(* IEC 61131-3 sources: veristc/veri-stc/tests/compiler-tests/negative, 18 files *)

(* ---- in_out_expr.st ---- *)
(* ================================================================
   negative/in_out_expr.st  --  VAR_IN_OUT 实参必须是简单变量名

   别名需要一个稳定的存储位置，表达式/常量没有地址可取，
   故 a1.ACC := SHARED + 1 必须被拒绝。
   ================================================================ *)

VAR_GLOBAL
  SHARED : DINT;
  a1 : ACCUM;
END_VAR

FUNCTION_BLOCK ACCUM
VAR_IN_OUT
  ACC : DINT;
END_VAR
  ACC := ACC + 1;
END_FUNCTION_BLOCK

PROGRAM MAIN
  a1(ACC := SHARED + 1);
END_PROGRAM

(* ---- in_out_local.st ---- *)
(* ================================================================
   negative/in_out_local.st  --  VAR_IN_OUT 别名目标不能是调用方局部

   MAIN 的 tick 是帧局部槽位（不在可寻址线性内存中），取不到地址，
   因此不能作为 a1.ACC 的别名目标。检查层必须以 alias 诊断拒绝。
   ================================================================ *)

VAR_GLOBAL
  a1 : ACCUM;
END_VAR

FUNCTION_BLOCK ACCUM
VAR_IN_OUT
  ACC : DINT;
END_VAR
  ACC := ACC + 1;
END_FUNCTION_BLOCK

PROGRAM MAIN
VAR
  tick : DINT;
END_VAR
  a1(ACC := tick);
END_PROGRAM

(* ---- in_out_type.st ---- *)
(* ================================================================
   negative/in_out_type.st  --  VAR_IN_OUT 两侧类型必须完全一致

   别名不经过隐式转换（同一块存储被两侧按同一宽度读写），
   且解引用指令按 4 字节定宽访问，故 INT(16 位) 目标必须拒绝。
   ================================================================ *)

VAR_GLOBAL
  SMALL : INT;
  a1 : ACCUM;
END_VAR

FUNCTION_BLOCK ACCUM
VAR_IN_OUT
  ACC : DINT;
END_VAR
  ACC := ACC + 1;
END_FUNCTION_BLOCK

PROGRAM MAIN
  a1(ACC := SMALL);
END_PROGRAM

(* ---- in_out_unbound.st ---- *)
(* ================================================================
   negative/in_out_unbound.st  --  VAR_IN_OUT 端口必须被绑定

   端口不绑定就没有别名目标（既无初值可拷贝，也无副本语义可言），
   与 IEC 要求一致：必须显式绑定到调用方存储。
   ================================================================ *)

VAR_GLOBAL
  SHARED : DINT;
  a1 : ACCUM;
END_VAR

FUNCTION_BLOCK ACCUM
VAR_IN_OUT
  ACC : DINT;
END_VAR
  ACC := ACC + 1;
END_FUNCTION_BLOCK

PROGRAM MAIN
  a1();
END_PROGRAM

(* ---- in_out_unknown_port.st ---- *)
(* ================================================================
   negative/in_out_unknown_port.st  --  调用只能绑定已声明端口

   FB_ACC 只声明了 ACC，调用点写 NOPE := SHARED 属于拼写/绕过声明，
   在逐引用端口上尤其危险（会把地址压进错误的槽位）。
   ================================================================ *)

VAR_GLOBAL
  SHARED : DINT;
  a1 : FB_ACC;
END_VAR

FUNCTION_BLOCK FB_ACC
VAR_IN_OUT
  ACC : DINT;
END_VAR
  ACC := ACC + 1;
END_FUNCTION_BLOCK

PROGRAM MAIN
  a1(ACC := SHARED, NOPE := SHARED);
END_PROGRAM

(* ---- literal_derived_name.st ---- *)
(* ================================================================
   negative/literal_derived_name.st -- 派生名不可书写

   expand_instances 产出的扁平全局名形如 a1#Q（'#' 为保留分隔符）。
   标识符文法是 字母 (字母|数字|_)*，不含 '#' ⇒ 源码里写 a1#Q 只能
   在词法阶段失败，用户无法伪造出一个"看起来像派生名"的名字去和
   真实派生名抢同一槽位，也不必再靠命名约定避免 a1_Q 这类碰撞。

   合法的字段访问写法是 IEC 点号 a1.Q，由 parser 融合为 a1#Q。
   ================================================================ *)

VAR_GLOBAL
  a1 : LATCH;
  x : DINT;
END_VAR

FUNCTION_BLOCK LATCH
VAR_OUTPUT
  Q : DINT;
END_VAR
  Q := 1;
END_FUNCTION_BLOCK

PROGRAM MAIN
  x := a1#Q;
END_PROGRAM

(* ---- name_collision_expanded.st ---- *)
(* ================================================================
   negative/name_collision_expanded.st -- 展开后派生名重复

   expand_instances（function_check.v）为实例 a1 的每个可写字段生成
   扁平全局名 a1#<字段>。若同一个 FUNCTION_BLOCK 里两个可写字段同名
   （此处 VAR_OUTPUT Q 与实例状态 VAR Q 重名），展开后就会产出两条
   a1#Q 声明 ⇒ 两个逻辑变量落到同一全局槽位、互相覆盖。

   这类冲突只在 prepare_program 之后才存在，因此 GATE-1 的重复名检查
   必须在展开后再跑一次，由 duplicate_declaration_msg 报出冲突的名字。

   （分隔符已改为标识符文法外的 '#'，用户无法手写派生名，所以静态
     命名冲突只剩"展开自身产出重名"这一条路径 —— 正是本用例。）
   ================================================================ *)

VAR_GLOBAL
  a1 : LATCH;
END_VAR

FUNCTION_BLOCK LATCH
VAR_INPUT
  K : DINT;
END_VAR
VAR_OUTPUT
  Q : DINT;
END_VAR
VAR
  Q : DINT;
END_VAR
  Q := K;
END_FUNCTION_BLOCK

PROGRAM MAIN
VAR
  tick : DINT;
END_VAR
  tick := CycleCounter();
  a1(K := tick);
END_PROGRAM

(* ---- qualified_in_out_read.st ---- *)
(* ================================================================
   negative/qualified_in_out_read.st -- 封装：别名端口不可用点号引用

   6.5.1 方向表的 VAR_IN_OUT 行。v1.5 起 VAR_IN_OUT 降级为"持有调用方
   存储地址的形参槽"（I32_LOAD_PTR / I32_STORE_PTR），expand_instances
   不为它生成派生全局，所以 `x := a1.ACC;` 引用的名字根本不存在，由类型
   检查阶段以 KIND=type 拒绝。

   这不是多余的严格性：调用方本来就持有别名目标（此处 shared），要读就
   直接读它 —— 读得到同一份存储，且不需要绕过 FB 的端口约定。

   与 qualified_input_read.st 的区别只在端口方向（IN_OUT vs INPUT）；
   与 qualified_internal_read.st（KIND=access）的区别在于名字是否存在。
   ================================================================ *)

(* 实例声明必须先于 POU 列表（顶层文法：VAR_GLOBAL → POU*）*)
VAR_GLOBAL
  a1 : ACCUM;
  shared : DINT;
  x : DINT;
END_VAR

FUNCTION_BLOCK ACCUM
VAR_INPUT
  K : DINT;
END_VAR
VAR_OUTPUT
  LAST : DINT;
END_VAR
VAR_IN_OUT
  ACC : DINT;
END_VAR
  LAST := ACC;
  ACC := ACC + K;
END_FUNCTION_BLOCK

PROGRAM MAIN
  a1(ACC := shared, K := 10);
  x := a1.ACC;
END_PROGRAM

(* ---- qualified_input_read.st ---- *)
(* ================================================================
   negative/qualified_input_read.st -- 封装：输入/别名端口不可用点号引用

   spec/safest-spec.md 6.5.1 方向表里 `VAR_INPUT` 与 `VAR_IN_OUT` 两行的
   体外访问都落到 `KIND=type`：expand_instances 只为可写字段
   （VAR_OUTPUT + 实例内 VAR）生成扁平派生全局，输入端口经调用点绑定为
   形参、别名端口降级为指针形参，二者都不存在名为 a1#K / a1#ACC 的全局。
   于是引用它们 = 引用未声明名，由类型检查阶段以 KIND=type 拒绝（而非
   access）。已知精度取舍：这条路径复用通用类型错误，诊断形如
     POU=MAIN VAR=- KIND=type LOC=- MSG=type error
   不指认具体名字，且报出第一条即中止（Fatal error）。因此本文件只保留
   一处违规（VAR_INPUT）；VAR_IN_OUT 的同一路径见 qualified_in_out_read.st，
   两行方向规则各自独立可验证。

   对比 qualified_internal_read.st（VAR=a1#C KIND=access）：那条是名字
   确实存在（内部 VAR 生成了派生全局）但封装禁止体外访问；本条是名字
   不存在。两者共同构成 6.5.1 方向表的机器可验证部分。
   ================================================================ *)

(* 实例声明必须先于 POU 列表（顶层文法：VAR_GLOBAL → POU*）*)
VAR_GLOBAL
  a1 : ACCUM;
  shared : DINT;
  x : DINT;
END_VAR

FUNCTION_BLOCK ACCUM
VAR_INPUT
  K : DINT;
END_VAR
VAR_OUTPUT
  LAST : DINT;
END_VAR
VAR_IN_OUT
  ACC : DINT;
END_VAR
  LAST := ACC;
  ACC := ACC + K;
END_FUNCTION_BLOCK

PROGRAM MAIN
  a1(ACC := shared, K := 10);
  x := a1.K;
END_PROGRAM

(* ---- qualified_internal_read.st ---- *)
(* ================================================================
   negative/qualified_internal_read.st -- 封装：内部状态对外不可见

   FB 的 VAR（实例持久状态，此处 C）是 FUNCTION_BLOCK 的私有内容：
   外部只能经 VAR_OUTPUT / VAR_IN_OUT 观察和交互。写 a1.C 会让调用方
   绕过 FB 的算法直接读内部计数器，多实例/维护场景下等价于破坏封装。

   expand_instances 本就不为 D_INPUT/D_IN_OUT 生成全局，但会为内部 VAR
   生成可写的扁平全局（FB 体内要读写它）；因此"外部不得引用"必须由
   访问规则单独把关 —— 诊断 KIND=access，VAR=a1#C 指认被泄漏的字段。
   ================================================================ *)

VAR_GLOBAL
  a1 : LATCH;
  x : DINT;
END_VAR

FUNCTION_BLOCK LATCH
VAR_INPUT
  K : DINT;
END_VAR
VAR_OUTPUT
  Q : DINT;
END_VAR
VAR
  C : DINT;
END_VAR
  C := C + 1;
  Q := K;
END_FUNCTION_BLOCK

PROGRAM MAIN
  a1(K := 3);
  x := a1.C;
END_PROGRAM

(* ---- qualified_output_write.st ---- *)
(* ================================================================
   negative/qualified_output_write.st -- 封装：输出只能由 FB 体写

   VAR_OUTPUT 是 FB 对外的只读结果。外部写 a1.Q 会在 FB 下一次执行之前
   篡改其结论，使"输出由算法决定"这条安全论证失效（同理 VAR_INPUT 由
   调用点绑定，也不能在体外的表达式里直接读写）。

   检查在 prepare_program 之后进行（派生名此时才存在），诊断 KIND=access
   并以 VAR=a1#Q 指认被篡改的字段。
   ================================================================ *)

VAR_GLOBAL
  a1 : LATCH;
END_VAR

FUNCTION_BLOCK LATCH
VAR_INPUT
  K : DINT;
END_VAR
VAR_OUTPUT
  Q : DINT;
END_VAR
  Q := K;
END_FUNCTION_BLOCK

PROGRAM MAIN
  a1(K := 3);
  a1.Q := 99;
END_PROGRAM

(* ---- iomap_unbound_name.st ---- *)
(* ================================================================
   negative/iomap_unbound_name.st -- IOMAP must bind a declared global

   An IOMAP entry names a global variable and gives it a physical channel.
   The compiler resolves that name to the variable's real global slot
   (build_global_env); a name that is not a declared global has no slot, so
   the entry could never be filled by the runtime. Accepting it would
   silently produce a program whose I/O quietly goes nowhere.

   Rejection: KIND=declaration, VAR=<the bad name>. Only the unbound entry
   is reported -- the well-formed one passes untouched.
   ================================================================ *)

VAR_GLOBAL
  ao0 : DINT;
END_VAR
IOMAP
  ao0, 1, OUTPUT, DINT;
  ghost, 2, INPUT, DINT;
END_IOMAP
PROGRAM P
  ao0 := 5;
END_PROGRAM

(* ---- real_literal_exponent.st ---- *)
(* Negative test: a REAL literal whose exponent leaves the exactness premises
   of the decimal-to-binary64 fast path.

   lexer.v scales a literal by a single power of ten that must itself be exactly
   representable: `E+n` needs significant digits + n <= 15, `E-n` needs fraction
   digits + n <= 22. 1.0e30 would require 10^30 (> 2^53), so it is refused
   (exit 21) rather than rounded twice. *)

PROGRAM real_literal_exponent
VAR
  x : REAL;
END_VAR
  x := 1.0e30;
END_PROGRAM

(* ---- real_literal_precision.st ---- *)
(* Negative test: a REAL literal with more significant digits than the
   decimal-to-binary64 fast path can produce exactly.

   lexer.v builds a real literal as mant / 10^k with both terms exactly
   representable, which needs at most 15 significant digits. A longer literal
   would need a second rounding step, so it is refused as a lexical failure
   (exit 21) instead of being silently double-rounded. *)

PROGRAM real_literal_precision
VAR
  x : REAL;
END_VAR
  x := 0.1234567890123456;
END_PROGRAM

(* ---- scope_violation.st ---- *)
(* Negative test: undeclared variable.
   Variable 'y' is never declared, so this must be rejected. *)

PROGRAM scope_violation
VAR
  x : DINT;
END_VAR
  x := y;
END_PROGRAM

(* ---- syntax_error.st ---- *)
(* Negative test: syntax error.
   Missing END_VAR causes a parse failure. *)

PROGRAM syntax_error
VAR
  x : DINT;
  x := 1;
END_PROGRAM

(* ---- type_mismatch.st ---- *)
(* Negative test: type mismatch.
   Assigning a BOOL value to a DINT variable is not allowed. *)

PROGRAM type_mismatch
VAR
  x : DINT;
  b : BOOL;
END_VAR
  b := TRUE;
  x := b;
END_PROGRAM

(* ---- uninit_var.st ---- *)
(* Negative test: FUNCTION modifies VAR_INPUT (purity violation).
   A FUNCTION must not assign to its input parameters. *)

FUNCTION Bad : DINT
VAR_INPUT
  x : DINT;
END_VAR
  x := 1;
  Bad := x;
END_FUNCTION

PROGRAM dup_main
VAR
  y : DINT;
END_VAR
  y := Bad(0);
END_PROGRAM
